(* IEC 61131-3 sources: iiot-demo/pous/programs, 1 file *)

(* ---- temp_check.st ---- *)
PROGRAM temp_check
  VAR
    rTemp : REAL;
    xAlarm : BOOL;
  END_VAR

xAlarm := rTemp > 80.0;

END_PROGRAM
